Fanuc KAREL source: kb00026.compact.KL

PROGRAM KB00026
%STACKSIZE=65535
%PRIORITY=65535
%NOLOCKGROUP
%ENVIRONMENT REGOPE
VAR
P1 : INTEGER
P2 : INTEGER
P3 : INTEGER
BEGIN
P1=1
P2=1
P3=1
CLR_POS_REG(P1,P2,P3)
END KB00026
